// TIA Portal project "项目6" (V15.1)

(* hardware
DEVICE "HMI_1"  KTP700 Basic PN
   slot 0: "HMI_1"  KTP700 Basic PN  6AV2 123-2GB03-0AX0  15.1.0.0
   slot 1: "HMI_RT_1"  KTP700 Basic PN  6AV2 123-2GB03-0AX0  15.1.0.0
   slot 5: "HMI_1.IE_CP_1"  PROFINET Interface  15.0.1.0
      slot 1: "PROFINET Interface_1"  PROFINET Interface
         slot 1: "Port_1"  Port
DEVICE "S7-1200 station_1"  S7-1200 Station
   slot 0: "Rack_0"  S7-1200 Rack  Rack  V1.0
   slot 1: "PLC_1"  CPU 1214C DC/DC/DC  6ES7 214-1AG40-0XB0  V4.2
   slot 2: "DI 16/DQ 16x24VDC_1"  6ES7 223-1BL32-0XB0  V2.0
   slot 3: "AI 4x13BIT/AQ 2x14BIT_1"  6ES7 234-4HE32-0XB0  V2.0
*)

// ===== PLC "PLC_1"  CPU 1214C DC/DC/DC =====

VAR_GLOBAL   // PLC tag table "默认变量表"
   "温度输入" AT %IW116 : Int;
   "灯开关" AT %I0.0 : Bool;
   "风扇" AT %Q9.6 : Bool;
   "灯" AT %Q0.0 : Bool;
   "风扇开关" AT %I0.1 : Bool;
   "PWM输出" AT %Q9.7 : Bool;
   "风扇启动指示灯" AT %Q0.1 : Bool;
   "KP" AT %QD12 : Real;
   "KI" AT %QD16 : Real;
   "输入控制上限" AT %QD20 : Real;
   "输入控制下限" AT %QD24 : Real;
   "当前偏差" AT %QD28 : Real;
   "上次偏差" AT %QD36 : Real;
   "当前温度值" AT %MD20 : Real;
   "PWM标志位" AT %QW44 : UInt;
   "PID输出值" AT %QD40 : Real;
   "目标占空比" AT %QW46 : Int;
   "PID增量" AT %QD48 : Real;
   "System_Byte" AT %MB1 : Byte;
   "FirstScan" AT %M1.0 : Bool;
   "DiagStatusUpdate" AT %M1.1 : Bool;
   "AlwaysTRUE" AT %M1.2 : Bool;
   "AlwaysFALSE" AT %M1.3 : Bool;
   "Clock_Byte" AT %MB0 : Byte;
   "Clock_10Hz" AT %M0.0 : Bool;
   "Clock_5Hz" AT %M0.1 : Bool;
   "Clock_2.5Hz" AT %M0.2 : Bool;
   "Clock_2Hz" AT %M0.3 : Bool;
   "Clock_1.25Hz" AT %M0.4 : Bool;
   "Clock_1Hz" AT %M0.5 : Bool;
   "Clock_0.625Hz" AT %M0.6 : Bool;
   "Clock_0.5Hz" AT %M0.7 : Bool;
END_VAR

DATA_BLOCK "PID数据"   // DB2
{ S7_Optimized_Access := 'TRUE' }
VERSION : 0.1
   VAR RETAIN
      设定值 : Real;
      模式选择 : Int;
   END_VAR
BEGIN
END_DATA_BLOCK

// folder: System blocks/Program resources

DATA_BLOCK "PLC_1_Send_DB"   // DB5
{ S7_Optimized_Access := 'TRUE' }
AUTHOR : SIMATIC
FAMILY : MC7Plus
NAME : TC_IP_v4
VERSION : 1.0
// stored: InstanceOfName TCON_IP_v4
"TCON_IP_v4"
BEGIN
   ID := 1;
   InterfaceId := 64;
   LocalPort := 2001;
END_DATA_BLOCK

// folder: (top level)

ORGANIZATION_BLOCK "Main"   // OB1, LAD, ProgramCycle
TITLE = "Main Program Sweep (Cycle)"
{ S7_Optimized_Access := 'TRUE' }
VERSION : 0.1
   VAR_INPUT
      Initial_Call : Bool;   // Initial call of this OB
      Remanence : Bool;   // =True, if remanent data are available
   END_VAR
BEGIN

REGION Network 1
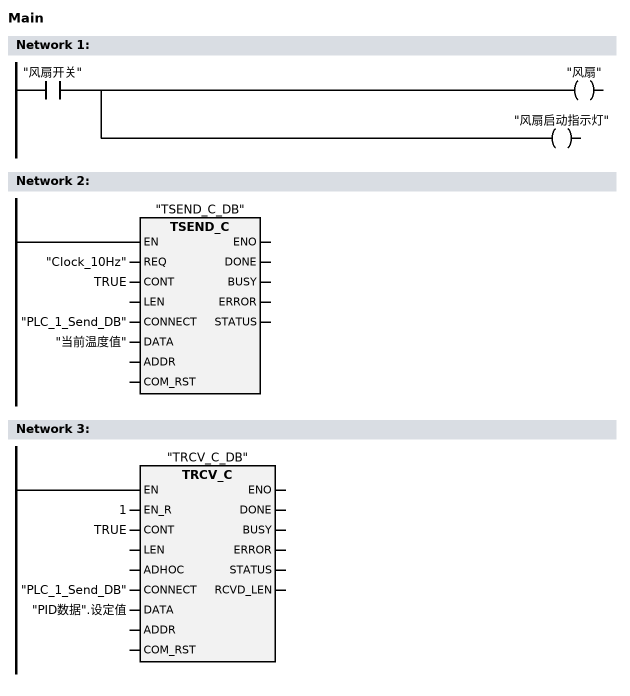
   RUNG wire#powerrail
      Contact( "风扇开关" )
      wire#w1
      Coil( "风扇" )
   END_RUNG
   RUNG wire#w1
      Coil( "风扇启动指示灯" )
   END_RUNG
   // the same network as SCL:
   "风扇" := "风扇开关";
   "风扇启动指示灯" := "风扇开关";
END_REGION

REGION Network 2
   "TSEND_C_DB"(REQ := "Clock_10Hz", CONT := TRUE, CONNECT := "PLC_1_Send_DB", DATA := "当前温度值");   // TSEND_C
END_REGION

REGION Network 3
   "TRCV_C_DB"(EN_R := 1, CONT := TRUE, CONNECT := "PLC_1_Send_DB", DATA := "PID数据".设定值);   // TRCV_C
END_REGION
END_ORGANIZATION_BLOCK

ORGANIZATION_BLOCK "Cyclic interrupt"   // OB30, SCL, CyclicInterrupt
{ S7_Optimized_Access := 'TRUE' }
VERSION : 0.1
   VAR_INPUT
      Initial_Call : Bool;   // Initial call of this OB
      Event_Count : Int;   // Events discarded
   END_VAR
BEGIN
   "当前温度值" := "温度输入" * 0.00361;
   "当前偏差" := "PID数据".设定值 - "当前温度值";
   "PID增量" := "KP" * ("当前偏差"-"上次偏差") +"KI" * "当前偏差";
   "PID输出值" := "PID输出值" + "PID增量";
   "上次偏差" := "当前偏差";
   IF "PID输出值" > 100 THEN
       // Statement section IF
       "PID输出值" := 100;
   END_IF;
   IF "PID输出值" < 0 THEN
       // Statement section IF
       "PID输出值" := 0;
   END_IF;

   "目标占空比" := REAL_TO_INT("PID输出值");
END_ORGANIZATION_BLOCK

ORGANIZATION_BLOCK "PWM输出程序"   // OB31, SCL, CyclicInterrupt
{ S7_Optimized_Access := 'TRUE' }
VERSION : 0.1
   VAR_INPUT
      Initial_Call : Bool;   // Initial call of this OB
      Event_Count : Int;   // Events discarded
   END_VAR
BEGIN
   "PWM标志位" := "PWM标志位" + 1;

   IF "PWM标志位" >= 100 THEN
       // Statement section IF
       "PWM标志位" := 0;
   END_IF;

   IF "PWM标志位" >= "目标占空比" THEN
       // Statement section IF
       "PWM输出" := 0;
   ELSE
       "PWM输出" := 1;
   END_IF;
END_ORGANIZATION_BLOCK

ORGANIZATION_BLOCK "Startup"   // OB100, SCL, Startup
TITLE = "Complete Restart"
{ S7_Optimized_Access := 'TRUE' }
VERSION : 0.1
   VAR_INPUT
      LostRetentive : Bool;   // True if retentive data are lost
      LostRTC : Bool;   // True if date and time are lost
   END_VAR
BEGIN
   "PID数据".设定值 := 45;
   "KP" := 12;
   "KI" := 0.2;
   "PWM标志位" := 0;
END_ORGANIZATION_BLOCK

(* ===== HMI "HMI_RT_1" =====
system functions are stored by id; their names below are inferred from use
connection "HMI_连接_1": ETHERNET, SMART_S7_1200_OMS

HMI tags "默认变量表"
   "Tag_ScreenNumber" : UInt, internal
   "PID数据_设定值" : Real = PLC PID数据.设定值, 1 s
   "KP" : Real = PLC KP AT %QD12, 1 s
   "KI" : Real = PLC KI AT %QD16, 1 s
   "PID输出值" : Real = PLC PID输出值 AT %QD40, 1 s
   "温度值" : Real = PLC 当前温度值 AT %MD20, 1 s

Template "模板_1" 800x480
   Button "退出" at 714,429 size 71x50; TextOff '退出'; PictureOff "ExitRuntime_KTP700_Basic_PN_TR"; PictureOn "ExitRuntime_KTP700_Basic_PN_TR"
      on Release: StopRuntime(0)
   Button "Template_Button" at 614,429 size 71x50; TextOff 'Text'
   Button "Template_Button_1" at 514,429 size 71x50; TextOff 'Text'
   Button "Template_Button_2" at 414,429 size 71x50; TextOff 'Text'
   Button "Template_Button_3" at 314,429 size 71x50; TextOff 'Text'
   Button "Template_Button_4" at 214,429 size 71x50; TextOff 'Text'
   Button "报警" at 114,429 size 71x50; TextOff '报警'; PictureOff "AlarmDisplay_KTP700_Basic_PN_TR"; PictureOn "AlarmDisplay_KTP700_Basic_PN_TR"
      on Release: function_ef3f5d25("报警窗口_Unacknowledged", -1)
   Button "起始画面" at 14,429 size 71x50; TextOff '起始画面'; PictureOff "NavigateHome_KTP700_Basic_PN_TR"; PictureOn "NavigateHome_KTP700_Basic_PN_TR"
      on Release: ActivateScreen("根画面", 0)
   SymbolicIOField "Symbolic_IO_Field_Screen" at 93,9 size 600x33; TextOff '0'; TextOn '1'; TextList "TextList_ScreenNames"
      ProcessValue <- "Tag_ScreenNumber"
      on Change: ActivateScreenByNumber("Tag_ScreenNumber", 0)
   DateTimeField "HmiScreenItemData" at 695,25 size 105x25
   DateTimeField "HmiScreenItemData_1" at 695,0 size 105x25
   GraphicView "Logo" at 0,0 size 91x51; Picture "HMI_1 的 Logo"

screen "根画面" 800x480, template "模板_1"
   on GenerateScreen: SetTag("Tag_ScreenNumber", 1)
   IOField "I/O 域_1" at 37,77 size 96x50; FormatPattern s99.99
      ProcessValue <- "PID数据_设定值"
   IOField "I/O 域_2" at 37,219 size 96x49; FormatPattern s99.99
      ProcessValue <- "KP"
   TrendView "趋势视图_1" at 183,57 size 600x358
   TextField "文本域_1" at 35,199 size 23x20; Text 'KP'
   TextField "文本域_2" at 37,57 size 90x20; Text '温度设定值'
   TextField "文本域_3" at 36,268 size 23x20; Text 'KI'
   IOField "I/O 域_3" at 36,289 size 96x51; FormatPattern s99.99
      ProcessValue <- "KI"
   TextField "文本域_4" at 34,127 size 56x20; Text '当前值'
   IOField "I/O 域_4" at 37,150 size 96x49; FormatPattern s99.99
      ProcessValue <- "温度值"
*)